Fanuc KAREL source: kb00107.compact.KL

PROGRAM KB00107
%STACKSIZE=65535
%PRIORITY=65535
%NOLOCKGROUP
VAR
P1 : XYZWPREXT
RESULT : BOOLEAN
BEGIN
RESULT=IN_RANGE(P1)
END KB00107
